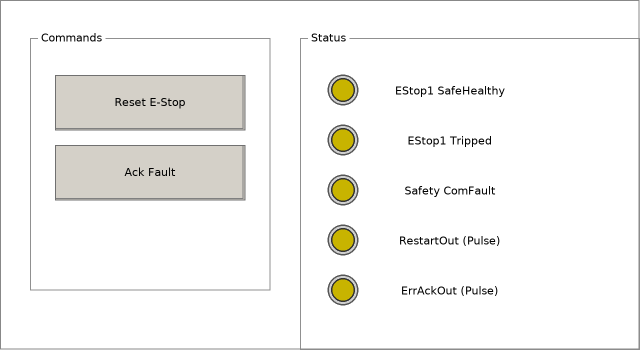
VISUALIZATION VISU_SafetySim  // 640x350
    GroupBox (300,30 340x320), "Status"
    GroupBox (30,30 240x260), "Commands"
    Lamp1 (325,72 36x36), variable: GVL_Safety.bEStop1_SafeHealthy, style: Lamp-Lamp1-Yellow
    Label (375,76 150x30), "EStop1 SafeHealthy"
    Label (375,176 150x30), "Safety ComFault"
    Label (375,126 150x30), "EStop1 Tripped"
    Label (375,276 150x30), "ErrAckOut (Pulse)"
    Label (375,226 150x30), "RestartOut (Pulse)"
    Lamp1 (325,122 36x36), variable: GVL_Safety.bEStop1_Tripped, style: Lamp-Lamp1-Yellow
    Lamp1 (325,172 36x36), variable: GVL_Safety.bSafety_ComFault, style: Lamp-Lamp1-Yellow
    Lamp1 (325,272 36x36), variable: GVL_Safety.bSafety_ErrAckOut, style: Lamp-Lamp1-Yellow
    Lamp1 (325,222 36x36), variable: GVL_Safety.bEStop1_RestartOut, style: Lamp-Lamp1-Yellow
    Button (55,75 190x55), "Reset E-Stop", pressed state: GVL_Safety.bEStop1_ResetCmd
        tap GVL_Safety.bEStop1_ResetCmd
    Button (55,145 190x55), "Ack Fault", pressed state: GVL_Safety.bSafety_ErrAckCmd
        tap GVL_Safety.bSafety_ErrAckCmd
END_VISUALIZATION

(* stored: Version 1.1.0.1
   Visu VISU_SafetySim: Id {84056c83-e112-424c-8449-25cff16d0cd7} *)
